// TIA Portal V21 export
// export: Created 2026-11-21T13:31:41.9480563Z, ExportSetting WithDefaults, DisplayName Totally Integrated Automation Portal, DisplayVersion V21, DisplayName STEP 7 Professional, DisplayVersion V21, DisplayName STEP 7 Safety, DisplayVersion V21, DisplayName Tech WebApplication, DisplayVersion V21, DisplayName WinCC Basic/Comfort/Advanced, DisplayVersion V21, DisplayName WinCC Unified, DisplayVersion V21
DATA_BLOCK "LineDb"   // DB43
VERSION : 0.1
// stored: AssignedProDiagFB PlantDiag, AutoNumber true, DBAccessibleFromOPCUA true, DBAccessibleFromWebserver true, InstanceOfName Line, InstanceOfType FB
"Line"
   // VAR_INPUT
   //    command : Bool;
   // END_VAR
   // VAR_OUTPUT
   //    running : Bool;
   // END_VAR
   // VAR
   //    drive { S7_SetPoint := 'True'} : "Motor";
   // END_VAR
BEGIN
END_DATA_BLOCK
